(* IEC 61131-3 sources: volt/packages/volt-lsp-iec/test-corpus/pro2193/Device/Plc Logic/Application/99 Library/Function Blocks/Actuators/Actuator, 3 files *)

(* ---- IActuator.itf ---- *)
INTERFACE IActuator

// Maps the actuator to the physical output
METHOD PUBLIC Map : BOOL

END_METHOD

// Reset the output (=False)
METHOD PUBLIC Reset

END_METHOD

// Set the output (=True)
METHOD PUBLIC Set : BOOL

END_METHOD

// Set the output True or False
METHOD PUBLIC SetOrReset
VAR_INPUT
	xValue	: BOOL;
END_VAR

END_METHOD

END_INTERFACE

(* ---- ActuatorFB.pou ---- *)
// Basic FB to control an output. No manual control!
{attribute 'monitoring_display' := 'output'}
{attribute 'symbol' := 'none'}
FUNCTION_BLOCK PUBLIC ActuatorFB
IMPLEMENTS IActuator
VAR
	{attribute 'symbol' := 'read'}	output					: BOOL;
	MeasureOnTime			: ONTIME;
	TimeOfLastSwitch		: DT;
END_VAR

%LANGUAGE ST
Counters();

END_FUNCTION_BLOCK

METHOD PRIVATE Counters

%LANGUAGE FBD
%NETWORK
// Calculate the on-time and the number of switches of the output
MeasureOnTime(In := output);
%NETWORK
// On a rising edge of the output, save the current date/time
MOVE(EN := RISING(output), TimeSettings.dtNow, OUT => TimeOfLastSwitch);
END_METHOD

// Maps the actuator to the physical output
METHOD PUBLIC Map : BOOL

%LANGUAGE ST
Map := output;

END_METHOD

// Reset the output (=False)
METHOD PUBLIC Reset

%LANGUAGE ST
output := FALSE;
END_METHOD

// Set the output (=True)
METHOD PUBLIC Set : BOOL

%LANGUAGE ST
output := TRUE;
END_METHOD

// Set the output True or False
METHOD PUBLIC SetOrReset
VAR_INPUT
	xValue	: BOOL;
END_VAR

%LANGUAGE ST
output := xValue;
END_METHOD

(* ---- ActuatorWithManualControlFB.pou ---- *)
// Basic actuator with manual control enabled
{attribute 'monitoring_display' := 'Output.output'}
{attribute 'symbol' := 'none'}
FUNCTION_BLOCK PUBLIC ActuatorWithManualControlFB
EXTENDS ActuatorWithManualControl_BaseFB
IMPLEMENTS IActuator
VAR
	{attribute 'symbol' := 'read'}	Output					: ActuatorFB;
END_VAR

%LANGUAGE ST
SUPER^();

END_FUNCTION_BLOCK

METHOD PROTECTED ManualControl
VAR_INPUT
	minButtonPushed			: BOOL;		// Both the software button (on screen) and the hardware button (if attached)
	plusButtonPushed		: BOOL;		// Both the software button (on screen) and the hardware button (if attached)
END_VAR

%LANGUAGE ST
IF plusButtonPushed THEN
	Set();
END_IF

IF minButtonPushed THEN
	Reset();
END_IF

END_METHOD

// Maps the actuator to the physical output
METHOD PUBLIC Map : BOOL

%LANGUAGE ST
Map := Output.Map();

END_METHOD

// Reset the output (=False)
METHOD PUBLIC Reset

%LANGUAGE ST
Output.Reset();

END_METHOD

// Set the output (=True)
METHOD PUBLIC Set : BOOL

%LANGUAGE ST
Output.Set();

END_METHOD

// Set the output True or False
METHOD PUBLIC SetOrReset
VAR_INPUT
	xValue	: BOOL;
END_VAR

%LANGUAGE ST
Output.SetOrReset(xValue);

END_METHOD
